// TIA Portal V20 export
// export: Created 2026-10-20T12:44:57.3841535Z, ExportSetting WithDefaults, DisplayName Totally Integrated Automation Portal, DisplayVersion V20 Update 6, DisplayName TIA Portal Openness, DisplayVersion V20 Update 6, DisplayName TIA Portal Version Control Interface, DisplayVersion V20 Update 6, DisplayName SINAMICS Startdrive Advanced, DisplayVersion V20 SP1, DisplayName SINAMICS Startdrive G130, G150, S120, S150, SINAMICS MV, G220, S200, S210, DisplayVersion V20 SP1, DisplayName SINAMICS Startdrive G110M, G120, G120C, G120D, G120P, G115D, DisplayVersion V20 SP1, DisplayName STEP 7 Professional, DisplayVersion V20 Update 6, DisplayName STEP 7 Safety, DisplayVersion V20 Update 2, DisplayName WinCC Basic/Comfort/Advanced, DisplayVersion V20 Update 6, DisplayName WinCC Unified, DisplayVersion V20 Update 6
FUNCTION "CNV_Charge_Settings_FC" : Void   // FC42, SCL
{ S7_Optimized_Access := 'TRUE' }
VERSION : 0.1
// stored: AutoNumber true, IsIECCheckEnabled false, SetENOAutomatically false, UDAEnableTagReadback false
BEGIN
   CASE "CNV_System_Selected" OF
       1: //SYSTEM 1
           CASE "CNV_Level_Selected" OF
               1:
                   "PopUps_DB".Buffer_Cnv_Settings_1 := "Settings_DB".LCnv_Sys[1].Cnv_Level[1].Cnv1;
                   "PopUps_DB".ECnv_Settings := "Settings_DB".ECnv_Sys[1];
                   "PopUps_DB".Buffer_Cnv_Settings_2 := "Settings_DB".LCnv_Sys[1].Cnv_Level[1].Cnv2;
               2:
                   "PopUps_DB".Buffer_Cnv_Settings_1 := "Settings_DB".LCnv_Sys[1].Cnv_Level[2].Cnv1;
                   "PopUps_DB".ECnv_Settings := "Settings_DB".ECnv_Sys[1];
                   "PopUps_DB".Buffer_Cnv_Settings_2 := "Settings_DB".LCnv_Sys[1].Cnv_Level[2].Cnv2;
               3:
                   "PopUps_DB".Buffer_Cnv_Settings_1 := "Settings_DB".LCnv_Sys[1].Cnv_Level[3].Cnv1;
                   "PopUps_DB".ECnv_Settings := "Settings_DB".ECnv_Sys[1];
                   "PopUps_DB".Buffer_Cnv_Settings_2 := "Settings_DB".LCnv_Sys[1].Cnv_Level[3].Cnv2;
               4:
                   "PopUps_DB".Buffer_Cnv_Settings_1 := "Settings_DB".LCnv_Sys[1].Cnv_Level[4].Cnv1;
                   "PopUps_DB".ECnv_Settings := "Settings_DB".ECnv_Sys[1];
                   "PopUps_DB".Buffer_Cnv_Settings_2 := "Settings_DB".LCnv_Sys[1].Cnv_Level[4].Cnv2;
               5:
                   "PopUps_DB".Buffer_Cnv_Settings_1 := "Settings_DB".LCnv_Sys[1].Cnv_Level[5].Cnv1;
                   "PopUps_DB".ECnv_Settings := "Settings_DB".ECnv_Sys[1];
                   "PopUps_DB".Buffer_Cnv_Settings_2 := "Settings_DB".LCnv_Sys[1].Cnv_Level[5].Cnv2;
               6:
                   "PopUps_DB".Buffer_Cnv_Settings_1 := "Settings_DB".LCnv_Sys[1].Cnv_Level[6].Cnv1;
                   "PopUps_DB".ECnv_Settings := "Settings_DB".ECnv_Sys[1];
                   "PopUps_DB".Buffer_Cnv_Settings_2 := "Settings_DB".LCnv_Sys[1].Cnv_Level[6].Cnv2;
               7:
                   "PopUps_DB".Buffer_Cnv_Settings_1 := "Settings_DB".LCnv_Sys[1].Cnv_Level[7].Cnv1;
                   "PopUps_DB".ECnv_Settings := "Settings_DB".ECnv_Sys[1];
                   "PopUps_DB".Buffer_Cnv_Settings_2 := "Settings_DB".LCnv_Sys[1].Cnv_Level[7].Cnv2;
               8:
                   "PopUps_DB".Buffer_Cnv_Settings_1 := "Settings_DB".LCnv_Sys[1].Cnv_Level[8].Cnv1;
                   "PopUps_DB".ECnv_Settings := "Settings_DB".ECnv_Sys[1];
                   "PopUps_DB".Buffer_Cnv_Settings_2 := "Settings_DB".LCnv_Sys[1].Cnv_Level[8].Cnv2;
           END_CASE;
       2: //SYSTEM 2
           CASE "CNV_Level_Selected" OF
               1:
                   "PopUps_DB".Buffer_Cnv_Settings_1 := "Settings_DB".LCnv_Sys[2].Cnv_Level[1].Cnv1;
                   "PopUps_DB".ECnv_Settings := "Settings_DB".ECnv_Sys[2];
                   "PopUps_DB".Buffer_Cnv_Settings_2 := "Settings_DB".LCnv_Sys[2].Cnv_Level[1].Cnv2;
               2:
                   "PopUps_DB".Buffer_Cnv_Settings_1 := "Settings_DB".LCnv_Sys[2].Cnv_Level[2].Cnv1;
                   "PopUps_DB".ECnv_Settings := "Settings_DB".ECnv_Sys[2];
                   "PopUps_DB".Buffer_Cnv_Settings_2 := "Settings_DB".LCnv_Sys[2].Cnv_Level[2].Cnv2;
               3:
                   "PopUps_DB".Buffer_Cnv_Settings_1 := "Settings_DB".LCnv_Sys[2].Cnv_Level[3].Cnv1;
                   "PopUps_DB".ECnv_Settings := "Settings_DB".ECnv_Sys[2];
                   "PopUps_DB".Buffer_Cnv_Settings_2 := "Settings_DB".LCnv_Sys[2].Cnv_Level[3].Cnv2;
               4:
                   "PopUps_DB".Buffer_Cnv_Settings_1 := "Settings_DB".LCnv_Sys[2].Cnv_Level[4].Cnv1;
                   "PopUps_DB".ECnv_Settings := "Settings_DB".ECnv_Sys[2];
                   "PopUps_DB".Buffer_Cnv_Settings_2 := "Settings_DB".LCnv_Sys[2].Cnv_Level[4].Cnv2;
               5:
                   "PopUps_DB".Buffer_Cnv_Settings_1 := "Settings_DB".LCnv_Sys[2].Cnv_Level[5].Cnv1;
                   "PopUps_DB".ECnv_Settings := "Settings_DB".ECnv_Sys[2];
                   "PopUps_DB".Buffer_Cnv_Settings_2 := "Settings_DB".LCnv_Sys[2].Cnv_Level[5].Cnv2;
               6:
                   "PopUps_DB".Buffer_Cnv_Settings_1 := "Settings_DB".LCnv_Sys[2].Cnv_Level[6].Cnv1;
                   "PopUps_DB".ECnv_Settings := "Settings_DB".ECnv_Sys[2];
                   "PopUps_DB".Buffer_Cnv_Settings_2 := "Settings_DB".LCnv_Sys[2].Cnv_Level[6].Cnv2;
               7:
                   "PopUps_DB".Buffer_Cnv_Settings_1 := "Settings_DB".LCnv_Sys[2].Cnv_Level[7].Cnv1;
                   "PopUps_DB".ECnv_Settings := "Settings_DB".ECnv_Sys[2];
                   "PopUps_DB".Buffer_Cnv_Settings_2 := "Settings_DB".LCnv_Sys[2].Cnv_Level[7].Cnv2;
               8:
                   "PopUps_DB".Buffer_Cnv_Settings_1 := "Settings_DB".LCnv_Sys[2].Cnv_Level[8].Cnv1;
                   "PopUps_DB".ECnv_Settings := "Settings_DB".ECnv_Sys[2];
                   "PopUps_DB".Buffer_Cnv_Settings_2 := "Settings_DB".LCnv_Sys[2].Cnv_Level[8].Cnv2;
           END_CASE;
       3: //SYSTEM 3
           CASE "CNV_Level_Selected" OF
               1:
                   "PopUps_DB".Buffer_Cnv_Settings_1 := "Settings_DB".LCnv_Sys[3].Cnv_Level[1].Cnv1;
                   "PopUps_DB".ECnv_Settings := "Settings_DB".ECnv_Sys[3];
                   "PopUps_DB".Buffer_Cnv_Settings_2 := "Settings_DB".LCnv_Sys[3].Cnv_Level[1].Cnv2;
               2:
                   "PopUps_DB".Buffer_Cnv_Settings_1 := "Settings_DB".LCnv_Sys[3].Cnv_Level[2].Cnv1;
                   "PopUps_DB".ECnv_Settings := "Settings_DB".ECnv_Sys[3];
                   "PopUps_DB".Buffer_Cnv_Settings_2 := "Settings_DB".LCnv_Sys[3].Cnv_Level[2].Cnv2;
               3:
                   "PopUps_DB".Buffer_Cnv_Settings_1 := "Settings_DB".LCnv_Sys[3].Cnv_Level[3].Cnv1;
                   "PopUps_DB".ECnv_Settings := "Settings_DB".ECnv_Sys[3];
                   "PopUps_DB".Buffer_Cnv_Settings_2 := "Settings_DB".LCnv_Sys[3].Cnv_Level[3].Cnv2;
               4:
                   "PopUps_DB".Buffer_Cnv_Settings_1 := "Settings_DB".LCnv_Sys[3].Cnv_Level[4].Cnv1;
                   "PopUps_DB".ECnv_Settings := "Settings_DB".ECnv_Sys[3];
                   "PopUps_DB".Buffer_Cnv_Settings_2 := "Settings_DB".LCnv_Sys[3].Cnv_Level[4].Cnv2;
               5:
                   "PopUps_DB".Buffer_Cnv_Settings_1 := "Settings_DB".LCnv_Sys[3].Cnv_Level[5].Cnv1;
                   "PopUps_DB".ECnv_Settings := "Settings_DB".ECnv_Sys[3];
                   "PopUps_DB".Buffer_Cnv_Settings_2 := "Settings_DB".LCnv_Sys[3].Cnv_Level[5].Cnv2;
               6:
                   "PopUps_DB".Buffer_Cnv_Settings_1 := "Settings_DB".LCnv_Sys[3].Cnv_Level[6].Cnv1;
                   "PopUps_DB".ECnv_Settings := "Settings_DB".ECnv_Sys[3];
                   "PopUps_DB".Buffer_Cnv_Settings_2 := "Settings_DB".LCnv_Sys[3].Cnv_Level[6].Cnv2;
               7:
                   "PopUps_DB".Buffer_Cnv_Settings_1 := "Settings_DB".LCnv_Sys[3].Cnv_Level[7].Cnv1;
                   "PopUps_DB".ECnv_Settings := "Settings_DB".ECnv_Sys[3];
                   "PopUps_DB".Buffer_Cnv_Settings_2 := "Settings_DB".LCnv_Sys[3].Cnv_Level[7].Cnv2;
               8:
                   "PopUps_DB".Buffer_Cnv_Settings_1 := "Settings_DB".LCnv_Sys[3].Cnv_Level[8].Cnv1;
                   "PopUps_DB".ECnv_Settings := "Settings_DB".ECnv_Sys[3];
                   "PopUps_DB".Buffer_Cnv_Settings_2 := "Settings_DB".LCnv_Sys[3].Cnv_Level[8].Cnv2;
           END_CASE;
       4: //SYSTEM 4
           CASE "CNV_Level_Selected" OF
               1:
                   "PopUps_DB".Buffer_Cnv_Settings_1 := "Settings_DB".LCnv_Sys[4].Cnv_Level[1].Cnv1;
                   "PopUps_DB".ECnv_Settings := "Settings_DB".ECnv_Sys[4];
                   "PopUps_DB".Buffer_Cnv_Settings_2 := "Settings_DB".LCnv_Sys[4].Cnv_Level[1].Cnv2;
               2:
                   "PopUps_DB".Buffer_Cnv_Settings_1 := "Settings_DB".LCnv_Sys[4].Cnv_Level[2].Cnv1;
                   "PopUps_DB".ECnv_Settings := "Settings_DB".ECnv_Sys[4];
                   "PopUps_DB".Buffer_Cnv_Settings_2 := "Settings_DB".LCnv_Sys[4].Cnv_Level[2].Cnv2;
               3:
                   "PopUps_DB".Buffer_Cnv_Settings_1 := "Settings_DB".LCnv_Sys[4].Cnv_Level[3].Cnv1;
                   "PopUps_DB".ECnv_Settings := "Settings_DB".ECnv_Sys[4];
                   "PopUps_DB".Buffer_Cnv_Settings_2 := "Settings_DB".LCnv_Sys[4].Cnv_Level[3].Cnv2;
               4:
                   "PopUps_DB".Buffer_Cnv_Settings_1 := "Settings_DB".LCnv_Sys[4].Cnv_Level[4].Cnv1;
                   "PopUps_DB".ECnv_Settings := "Settings_DB".ECnv_Sys[4];
                   "PopUps_DB".Buffer_Cnv_Settings_2 := "Settings_DB".LCnv_Sys[4].Cnv_Level[4].Cnv2;
               5:
                   "PopUps_DB".Buffer_Cnv_Settings_1 := "Settings_DB".LCnv_Sys[4].Cnv_Level[5].Cnv1;
                   "PopUps_DB".ECnv_Settings := "Settings_DB".ECnv_Sys[4];
                   "PopUps_DB".Buffer_Cnv_Settings_2 := "Settings_DB".LCnv_Sys[4].Cnv_Level[5].Cnv2;
               6:
                   "PopUps_DB".Buffer_Cnv_Settings_1 := "Settings_DB".LCnv_Sys[4].Cnv_Level[6].Cnv1;
                   "PopUps_DB".ECnv_Settings := "Settings_DB".ECnv_Sys[4];
                   "PopUps_DB".Buffer_Cnv_Settings_2 := "Settings_DB".LCnv_Sys[4].Cnv_Level[6].Cnv2;
               7:
                   "PopUps_DB".Buffer_Cnv_Settings_1 := "Settings_DB".LCnv_Sys[4].Cnv_Level[7].Cnv1;
                   "PopUps_DB".ECnv_Settings := "Settings_DB".ECnv_Sys[4];
                   "PopUps_DB".Buffer_Cnv_Settings_2 := "Settings_DB".LCnv_Sys[4].Cnv_Level[7].Cnv2;
               8:
                   "PopUps_DB".Buffer_Cnv_Settings_1 := "Settings_DB".LCnv_Sys[4].Cnv_Level[8].Cnv1;
                   "PopUps_DB".ECnv_Settings := "Settings_DB".ECnv_Sys[4];
                   "PopUps_DB".Buffer_Cnv_Settings_2 := "Settings_DB".LCnv_Sys[4].Cnv_Level[8].Cnv2;
           END_CASE;
       5: //SYSTEM 5
           CASE "CNV_Level_Selected" OF
               1:
                   "PopUps_DB".Buffer_Cnv_Settings_1 := "Settings_DB".LCnv_Sys[5].Cnv_Level[1].Cnv1;
                   "PopUps_DB".ECnv_Settings := "Settings_DB".ECnv_Sys[5];
                   "PopUps_DB".Buffer_Cnv_Settings_2 := "Settings_DB".LCnv_Sys[5].Cnv_Level[1].Cnv2;
               2:
                   "PopUps_DB".Buffer_Cnv_Settings_1 := "Settings_DB".LCnv_Sys[5].Cnv_Level[2].Cnv1;
                   "PopUps_DB".ECnv_Settings := "Settings_DB".ECnv_Sys[5];
                   "PopUps_DB".Buffer_Cnv_Settings_2 := "Settings_DB".LCnv_Sys[5].Cnv_Level[2].Cnv2;
               3:
                   "PopUps_DB".Buffer_Cnv_Settings_1 := "Settings_DB".LCnv_Sys[5].Cnv_Level[3].Cnv1;
                   "PopUps_DB".ECnv_Settings := "Settings_DB".ECnv_Sys[5];
                   "PopUps_DB".Buffer_Cnv_Settings_2 := "Settings_DB".LCnv_Sys[5].Cnv_Level[3].Cnv2;
               4:
                   "PopUps_DB".Buffer_Cnv_Settings_1 := "Settings_DB".LCnv_Sys[5].Cnv_Level[4].Cnv1;
                   "PopUps_DB".ECnv_Settings := "Settings_DB".ECnv_Sys[5];
                   "PopUps_DB".Buffer_Cnv_Settings_2 := "Settings_DB".LCnv_Sys[5].Cnv_Level[4].Cnv2;
               5:
                   "PopUps_DB".Buffer_Cnv_Settings_1 := "Settings_DB".LCnv_Sys[5].Cnv_Level[5].Cnv1;
                   "PopUps_DB".ECnv_Settings := "Settings_DB".ECnv_Sys[5];
                   "PopUps_DB".Buffer_Cnv_Settings_2 := "Settings_DB".LCnv_Sys[5].Cnv_Level[5].Cnv2;
               6:
                   "PopUps_DB".Buffer_Cnv_Settings_1 := "Settings_DB".LCnv_Sys[5].Cnv_Level[6].Cnv1;
                   "PopUps_DB".ECnv_Settings := "Settings_DB".ECnv_Sys[5];
                   "PopUps_DB".Buffer_Cnv_Settings_2 := "Settings_DB".LCnv_Sys[5].Cnv_Level[6].Cnv2;
               7:
                   "PopUps_DB".Buffer_Cnv_Settings_1 := "Settings_DB".LCnv_Sys[5].Cnv_Level[7].Cnv1;
                   "PopUps_DB".ECnv_Settings := "Settings_DB".ECnv_Sys[5];
                   "PopUps_DB".Buffer_Cnv_Settings_2 := "Settings_DB".LCnv_Sys[5].Cnv_Level[7].Cnv2;
               8:
                   "PopUps_DB".Buffer_Cnv_Settings_1 := "Settings_DB".LCnv_Sys[5].Cnv_Level[8].Cnv1;
                   "PopUps_DB".ECnv_Settings := "Settings_DB".ECnv_Sys[5];
                   "PopUps_DB".Buffer_Cnv_Settings_2 := "Settings_DB".LCnv_Sys[5].Cnv_Level[8].Cnv2;
           END_CASE;
   END_CASE;
END_FUNCTION
